(* IEC 61131-3 sources: Elmo_Master/Lasal_PRG/Elmo_EtherCAT_Test_4Axis/Class/ECAT_Master_Base (part 3) *)

#ifdef ECAT_DEBUG_EVENT_CALLBACKS
      LogError("ECAT-DEBUG: Event ECATM_EVTC_DC_DISABLED occured");
#endif

//*******************************************************************************************************************************************************
    ECATM_EVTC_ESM_DC_FAILED:
    //Error code used as argument of the ECATM_EVTC_MST_TRANS_FAILED or ECATM_EVTC_SLV_TRANS_FAILED event after the DC module failed.

#ifdef ECAT_DEBUG_EVENT_CALLBACKS
      LogError("ECAT-DEBUG: Event ECATM_EVTC_ESM_DC_FAILED occured");
#endif

//*******************************************************************************************************************************************************
    ECATM_EVTC_EOE_MBX_BAD_RSP:
    //Invalid EoE mailbox size received
    //arg1 ... slave index: int
    //arg2 ... EoE mailbox size:
    //arg3 ... EoE mailbox frame type: int

#ifdef ECAT_DEBUG_EVENT_CALLBACKS
      LogValue("ECAT-DEBUG: Invalid EoE mailbox size received. SlaveIndex: 0x{0}",evt^.arg1$UDINT);
      LogValue("ECAT-DEBUG: MBxSize: 0x{0}, MBxFrameType: 0x{1}",evt^.arg2$UDINT, evt^.arg3$UDINT);
#endif

//*******************************************************************************************************************************************************
    ECATM_EVTC_EOE_FRM_TRF_TMO:
    //Frame fragment timeout occurred. Frame was dropped
    //arg1 ... slave index: int

#ifdef ECAT_DEBUG_EVENT_CALLBACKS
      LogValue("ECAT-DEBUG: Invalid EoE mailbox size received. SlaveIndex: 0x{0}",evt^.arg1$UDINT);
#endif

//*******************************************************************************************************************************************************
    ECATM_EVTC_EOE_FRM_DROP_HDL:
    //Frame dropped because of no free frame handle available
    //arg1 ... slave index: int

#ifdef ECAT_DEBUG_EVENT_CALLBACKS
      LogValue("ECAT-DEBUG: EOE: Frame dropped because of no free frame handle available. SlaveIndex: 0x{0}",evt^.arg1$UDINT);
#endif

//*******************************************************************************************************************************************************
    ECATM_EVTC_EOE_FRM_DROP_SIZE:
    //Frame with invalid size received. Frame was dropped
    //arg1 ... slave index: int

#ifdef ECAT_DEBUG_EVENT_CALLBACKS
      LogValue("ECAT-DEBUG: EOE: Frame with invalid size received. Frame was dropped. SlaveIndex: 0x{0}",evt^.arg1$UDINT);
#endif

//*******************************************************************************************************************************************************
    ECATM_EVTC_EOE_SAT_MAC_ADD:
    //Frame with a not yet known MAC received. MAC added to switch address table
    //arg1 ... Device index: int
    //arg2 ... arg3 MAC address: arg2[3] : arg2[2] : arg2[1] : arg2[0] : arg3[1] : arg2[0]

#ifdef ECAT_DEBUG_EVENT_CALLBACKS
      LogValue("ECAT-DEBUG: EOE: Frame with a not yet known MAC received. MAC added to switch address table. DeviceIndex: 0x{0}",evt^.arg1$UDINT);
      LogValue("ECAT-DEBUG: MACADDR: 0x{0}0x{1}",evt^.arg2$UDINT, evt^.arg3$UDINT);//Before Use, should be formated correctly
#endif

//*******************************************************************************************************************************************************
    ECATM_EVTC_EOE_SAT_MAC_RM:
    //MAC is dropped from switch address table
    //arg1 ... Device index: int
    //arg2 ... arg3 MAC address: arg2[3] : arg2[2] : arg2[1] : arg2[0] : arg3[1] : arg2[0]

#ifdef ECAT_DEBUG_EVENT_CALLBACKS
      LogValue("ECAT-DEBUG: EOE: MACAddr is dropped from switch address table. DeviceIndex: 0x{0}",evt^.arg1$UDINT);
      LogValue("ECAT-DEBUG: MACADDR: 0x{0}0x{1}",evt^.arg2$UDINT, evt^.arg3$UDINT);//Before Use, should be formated correctly
#endif

//*******************************************************************************************************************************************************
    ECATM_EVTC_FRM_BAD_FRMIDX:
    // A frame with a bad index was received
    // arg1 max allowed IDX field value: int
    // arg2 received IDX field value: int

#ifdef ECAT_DEBUG_EVENT_CALLBACKS
    HWC_LogPrintf(pThis:=this, format:="@ECAT-DEBUG: A frame with a bad index was received");
    HWC_LogPrintf(pThis:=this, format:="@ECAT-DEBUG: max allowed IDX field value: %d received IDX field value: %d.", #evt^.arg1, #evt^.arg2);
#endif

//*******************************************************************************************************************************************************
    ECATM_EVTC_FRM_CFG_OP_SIZE:
    // maximal frame size during OP is too small
    // arg1 configured value (_ecatm_cfg field frmsizeop): int
    // arg2 required value: int

#ifdef ECAT_DEBUG_EVENT_CALLBACKS
    HWC_LogPrintf(pThis:=this, format:="@ECAT-DEBUG: Maximal frame size during OP is too small");
    HWC_LogPrintf(pThis:=this, format:="@ECAT-DEBUG: configured value (_ecatm_cfg field frmsizeop): %d required value: %d.", #evt^.arg1, #evt^.arg2);
#endif

//*******************************************************************************************************************************************************
    ECATM_EVTC_CRD_STATUS_CHANGED:
    // The status of the network cable redundancy diagnostics has changed
    // arg1 _ecatm_crd_status pos0 field: int
    // arg2 _ecatm_crd_status pos1 field: int
    // arg3 _ecatm_crd_status flags field: int

#ifdef ECAT_DEBUG_EVENT_CALLBACKS
    HWC_LogPrintf(pThis:=this, format:="@ECAT-DEBUG: The status of the network cable redundancy diagnostics has changed");
    HWC_LogPrintf(pThis:=this, format:="@ECAT-DEBUG: _ecatm_crd_status pos0 field: %d _ecatm_crd_status pos1 field: %d.", #evt^.arg1, #evt^.arg2);
    HWC_LogPrintf(pThis:=this, format:="@ECAT-DEBUG: _ecatm_crd_status flags field: %d", #evt^.arg3);
#endif

//*******************************************************************************************************************************************************
    ECATM_EVTC_SOE_SSC_NOTIFY:
    // SoE Notify received
    // arg1 slave index: int
    // arg2 driveno: uint8_t
    // arg3 idn: uint16_t
    // arg4 status data (16bit) from slave

#ifdef ECAT_DEBUG_EVENT_CALLBACKS
    HWC_LogPrintf(pThis:=this, format:="@ECAT-DEBUG: SoE Notify received");
    HWC_LogPrintf(pThis:=this, format:="@ECAT-DEBUG: slave index: %d driveno: uint8_t: %d.", #evt^.arg1, #evt^.arg2);
    HWC_LogPrintf(pThis:=this, format:="@ECAT-DEBUG: idn: %d status data (16bit) from slave: %d", #evt^.arg3, #evt^.arg4);
#endif

//*******************************************************************************************************************************************************
    ECATM_EVTC_SOE_SSC_TRF_TMO:
    // SoE timeout error detected
    // arg1

#ifdef ECAT_DEBUG_EVENT_CALLBACKS
    HWC_LogPrintf(pThis:=this, format:="@ECAT-DEBUG: SoE timeout error detected");
#endif

//*******************************************************************************************************************************************************
    ECATM_EVTC_SOE_SSC_TRF_ERR:
    // SoE slave responded with an error
    // arg1 slave index: int
    // arg2 driveno: uint8_t
    // arg3 idn: uint16_t
    // arg4 SoE error code from slave: uint16_t

#ifdef ECAT_DEBUG_EVENT_CALLBACKS
    HWC_LogPrintf(pThis:=this, format:="@ECAT-DEBUG: SoE slave responded with an error");
    HWC_LogPrintf(pThis:=this, format:="@ECAT-DEBUG: slave index: %d driveno: uint8_t: %d.", #evt^.arg1, #evt^.arg2);
    HWC_LogPrintf(pThis:=this, format:="@ECAT-DEBUG: idn: %d SoE error code from slave: uint16_t: %d", #evt^.arg3, #evt^.arg4);
#endif

//*******************************************************************************************************************************************************
    ECATM_EVTC_SOE_SSC_BAD_RSP:
    // Bad SoE response received
    // arg1 slave index: int

#ifdef ECAT_DEBUG_EVENT_CALLBACKS
    HWC_LogPrintf(pThis:=this, format:="@ECAT-DEBUG: Bad SoE response received. slave index: %d", #evt^.arg1);
#endif

//*******************************************************************************************************************************************************
    ECATM_EVTC_SOE_SSC_RD_BUFSIZE:
    // SoE read failed because of invalid receive buffer size
    // arg1 slave index: int
    // arg2 driveno: uint8_t
    // arg3 idn: uint16_t
    // arg4 required size: int

#ifdef ECAT_DEBUG_EVENT_CALLBACKS
    HWC_LogPrintf(pThis:=this, format:="@ECAT-DEBUG: SoE read failed because of invalid receive buffer size");
    HWC_LogPrintf(pThis:=this, format:="@ECAT-DEBUG: slave index: %d driveno: uint8_t: %d.", #evt^.arg1, #evt^.arg2);
    HWC_LogPrintf(pThis:=this, format:="@ECAT-DEBUG: idn: %d required size: %d", #evt^.arg3, #evt^.arg4);
#endif

//*******************************************************************************************************************************************************
    ECATM_EVTC_SOE_SSC_RD_FRAG:
    // SoE read failed because of unexpected fragment number
    // arg1 slave index: int
    // arg2 driveno: uint8_t
    // arg3 idn: uint16_t

#ifdef ECAT_DEBUG_EVENT_CALLBACKS
    HWC_LogPrintf(pThis:=this, format:="@ECAT-DEBUG: SoE read failed because of unexpected fragment number");
    HWC_LogPrintf(pThis:=this, format:="@ECAT-DEBUG: slave index: %d driveno: uint8_t: %d.", #evt^.arg1, #evt^.arg2);
    HWC_LogPrintf(pThis:=this, format:="@ECAT-DEBUG: idn: %d.", #evt^.arg3);
#endif

//*******************************************************************************************************************************************************
    ECATM_EVTC_SII_EEPROM_BUSY_TMO:
    // SII EEPROM access failed because of EEPROM busy flag
    // arg1 slave index: int
    // arg2 SII Status Register (ESC register 0x502): uint8_t

#ifdef ECAT_DEBUG_EVENT_CALLBACKS
    HWC_LogPrintf(pThis:=this, format:="@ECAT-DEBUG: SII EEPROM access failed because of EEPROM busy flag");
    HWC_LogPrintf(pThis:=this, format:="@ECAT-DEBUG: slave index: %d SII Status Register (ESC register 0x502): uint8_t: %x.", #evt^.arg1, #evt^.arg2);
#endif

//*******************************************************************************************************************************************************
    ECATM_EVTC_SII_EEPROM_PDI_TMO:
    // SII EEPROM access failed as owenership is with PDI
    // arg1 slave index: int

#ifdef ECAT_DEBUG_EVENT_CALLBACKS
    HWC_LogPrintf(pThis:=this, format:="@ECAT-DEBUG: SII EEPROM access failed as owenership is with PDI. slave index: %d", #evt^.arg1);
#endif

//*******************************************************************************************************************************************************
    ECATM_EVTC_SII_INVALID_VERSION:
    // SII read till end failed as SII version is invalid
    // arg1 slave index: int
    // arg2 SII version field (0x3F) (should be 0x001): uint16_t

#ifdef ECAT_DEBUG_EVENT_CALLBACKS
    HWC_LogPrintf(pThis:=this, format:="@ECAT-DEBUG: SII read till end failed as SII version is invalid");
    HWC_LogPrintf(pThis:=this, format:="@ECAT-DEBUG: slave index: %d SII version field (0x3F) (should be 0x001): %x.", #evt^.arg1, #evt^.arg2);
#endif

//*******************************************************************************************************************************************************
    ECATM_EVTC_HC_TOO_MANY_DEVICES:
    // The number of found devices during HC detection exceeds the number of devices defined in the ENI
    // arg1 found devices: int
    // arg2 number of devices in ENI: int

#ifdef ECAT_DEBUG_EVENT_CALLBACKS
    HWC_LogPrintf(pThis:=this, format:="@ECAT-DEBUG: The number of found devices during HC detection exceeds the number of devices defined in the ENI");
    HWC_LogPrintf(pThis:=this, format:="@ECAT-DEBUG: found devices: %d number of devices in ENI: %d.", #evt^.arg1, #evt^.arg2);
#endif

//*******************************************************************************************************************************************************
    ECATM_EVTC_HC_GRP_SEARCH:
    // Start searching for matching HC group connected to a device port
    // arg1 slave index: int
    // arg2 port index: enum {ECAT_ESC_PORT_A; ECAT_ESC_PORT_B; ECAT_ESC_PORT_C; ECAT_ESC_PORT_D}

#ifdef ECAT_DEBUG_EVENT_CALLBACKS
    HWC_LogPrintf(pThis:=this, format:="@ECAT-DEBUG: Start searching for matching HC group connected to a device port");
    HWC_LogPrintf(pThis:=this, format:="@ECAT-DEBUG: slave index: %d port index: %d.", #evt^.arg1, #evt^.arg2);
#endif

//*******************************************************************************************************************************************************
    ECATM_EVTC_HC_GRP_FOUND:
    // Found a matching HC group connected to the device port
    // arg1 HC group index matching: int
    // arg2 slave index: int
    // arg3 port index: enum {ECAT_ESC_PORT_A; ECAT_ESC_PORT_B; ECAT_ESC_PORT_C; ECAT_ESC_PORT_D}

#ifdef ECAT_DEBUG_EVENT_CALLBACKS
    HWC_LogPrintf(pThis:=this, format:="@ECAT-DEBUG: Found a matching HC group connected to the device port");
    HWC_LogPrintf(pThis:=this, format:="@ECAT-DEBUG: HC group index that is no longer reachable: %d.", #evt^.arg1);
    HWC_LogPrintf(pThis:=this, format:="@ECAT-DEBUG: slave index: %d port index: %d.", #evt^.arg2, #evt^.arg3);
#endif

//*******************************************************************************************************************************************************
    ECATM_EVTC_HC_GRP_NO_MATCH:
    // Failed to find a matching HC group for the device port
    // arg1 slave index: int
    // arg2 port index: enum {ECAT_ESC_PORT_A; ECAT_ESC_PORT_B; ECAT_ESC_PORT_C; ECAT_ESC_PORT_D}

#ifdef ECAT_DEBUG_EVENT_CALLBACKS
    HWC_LogPrintf(pThis:=this, format:="@ECAT-DEBUG: Failed to find a matching HC group for the device port");
    HWC_LogPrintf(pThis:=this, format:="@ECAT-DEBUG: slave index: %d port index: %d.", #evt^.arg1, #evt^.arg2);
#endif

//*******************************************************************************************************************************************************
    ECATM_EVTC_HC_GRP_DISCONNECTED:
    // Hot Connect group is disconnected from the device port
    // arg1 HC group index that is no longer reachable: int
    // arg2 slave index: int
    // arg3 port index: enum {ECAT_ESC_PORT_A; ECAT_ESC_PORT_B; ECAT_ESC_PORT_C; ECAT_ESC_PORT_D}

#ifdef ECAT_DEBUG_EVENT_CALLBACKS
    HWC_LogPrintf(pThis:=this, format:="@ECAT-DEBUG: Hot Connect group is disconnected from the device port");
    HWC_LogPrintf(pThis:=this, format:="@ECAT-DEBUG: HC group index that is no longer reachable: %d.", #evt^.arg1);
    HWC_LogPrintf(pThis:=this, format:="@ECAT-DEBUG: slave index: %d port index: %d.", #evt^.arg2, #evt^.arg3);
#endif

//*******************************************************************************************************************************************************
    ECATM_EVTC_HC_PORT_CHANGED:
    // The status of device port has changed
    // arg1 slave index: int
    // arg2 port index: enum {ECAT_ESC_PORT_A; ECAT_ESC_PORT_B; ECAT_ESC_PORT_C; ECAT_ESC_PORT_D}
    // arg3 new status: flags see ECATM_HC_PORT_FLAG…
    // arg4 old status: flags see ECATM_HC_PORT_FLAG…

#ifdef ECAT_DEBUG_EVENT_CALLBACKS
    HWC_LogPrintf(pThis:=this, format:="@ECAT-DEBUG: The status of device port has changed");
    HWC_LogPrintf(pThis:=this, format:="@ECAT-DEBUG: slave index: %d port index: %d.", #evt^.arg1, #evt^.arg2);
    HWC_LogPrintf(pThis:=this, format:="@ECAT-DEBUG: new status: %d old status: %d.", #evt^.arg3, #evt^.arg4);
#endif

//*******************************************************************************************************************************************************
    ECATM_EVTC_HC_PORT_OPEN:
    // A device port will be opened to connect new devices
    // arg1 slave index: int
    // arg2 port index: enum {ECAT_ESC_PORT_A; ECAT_ESC_PORT_B; ECAT_ESC_PORT_C; ECAT_ESC_PORT_D}

#ifdef ECAT_DEBUG_EVENT_CALLBACKS
    HWC_LogPrintf(pThis:=this, format:="@ECAT-DEBUG: A device port will be opened to connect new devices");
    HWC_LogPrintf(pThis:=this, format:="@ECAT-DEBUG: slave index: %d port index: %d.", #evt^.arg1, #evt^.arg2);
#endif

//*******************************************************************************************************************************************************
    ECATM_EVTC_HC_MAN_PORT_CLOSED:
    // A mandatory connection at the device port is closed/disconnected
    // arg1 slave index: int
    // arg2 port index: enum {ECAT_ESC_PORT_A; ECAT_ESC_PORT_B; ECAT_ESC_PORT_C; ECAT_ESC_PORT_D}

#ifdef ECAT_DEBUG_EVENT_CALLBACKS
    HWC_LogPrintf(pThis:=this, format:="@ECAT-DEBUG: A mandatory connection at the device port is closed/disconnected");
    HWC_LogPrintf(pThis:=this, format:="@ECAT-DEBUG: slave index: %d port index: %d.", #evt^.arg1, #evt^.arg2);
#endif

//*******************************************************************************************************************************************************
    ECATM_EVTC_HC_MAN_PORT_OPENING:
    // Opening a connection at the device port which is closed
    // arg1 slave index: int
    // arg2 port index: enum {ECAT_ESC_PORT_A; ECAT_ESC_PORT_B; ECAT_ESC_PORT_C; ECAT_ESC_PORT_D}

#ifdef ECAT_DEBUG_EVENT_CALLBACKS
    HWC_LogPrintf(pThis:=this, format:="@ECAT-DEBUG: Opening a connection at the device port which is closed");
    HWC_LogPrintf(pThis:=this, format:="@ECAT-DEBUG: slave index: %d port index: %d.", #evt^.arg1, #evt^.arg2);
#endif

//*******************************************************************************************************************************************************
    ECATM_EVTC_HC_TOPO_INVALID:
    // The Hot Connect topology solver failed to match the current network topology

#ifdef ECAT_DEBUG_EVENT_CALLBACKS
    HWC_LogPrintf(pThis:=this, format:="@ECAT-DEBUG: The Hot Connect topology solver failed to match the current network topology");
#endif

//*******************************************************************************************************************************************************
    ECATM_EVTC_HC_SLV_NOT_CONNECTED:
    // The current device is part of a not connected HC group

#ifdef ECAT_DEBUG_EVENT_CALLBACKS
    HWC_LogPrintf(pThis:=this, format:="@ECAT-DEBUG: The current device is part of a not connected HC group");
#endif

//*******************************************************************************************************************************************************
    ECATM_EVTC_DC_PROPDLY_UPDATE:
    // The Distributed Clocks module is starting an propagation delay update run
    // The force flag is set when not triggered via _ecatm_dc_cfg.propdly_update_ms timeout.
    // arg1 forced run: bool

#ifdef ECAT_DEBUG_EVENT_CALLBACKS
    HWC_LogPrintf(pThis:=this, format:="@ECAT-DEBUG: The Distributed Clocks module is starting an propagation delay update run");
    HWC_LogPrintf(pThis:=this, format:="@ECAT-DEBUG: The force flag is set when not triggered via _ecatm_dc_cfg.propdly_update_ms timeout. forced run: %d", #evt^.arg1);
#endif

//*******************************************************************************************************************************************************
    ECATM_EVTC_DC_PROPDLY_FINISHED:
    // The propagation delay is now updated

#ifdef ECAT_DEBUG_EVENT_CALLBACKS
    HWC_LogPrintf(pThis:=this, format:="@ECAT-DEBUG: The propagation delay is now updated");
#endif

//*******************************************************************************************************************************************************
    ECATM_EVTC_DC_SLV_SYNC_TIMOUT:
    // The static drift compensation for a single device during during operation failed
    // arg1 slave index: int
    // arg2 last syncwin measured: unsigned int

#ifdef ECAT_DEBUG_EVENT_CALLBACKS
    HWC_LogPrintf(pThis:=this, format:="@ECAT-DEBUG: The static drift compensation for a single device during during operation failed");
    HWC_LogPrintf(pThis:=this, format:="@ECAT-DEBUG: slave index: %d last syncwin measured: %d.", #evt^.arg1, #evt^.arg2);
#endif

//*******************************************************************************************************************************************************
    ECATM_EVTC_FOE_ERROR_RSP:
    // Error code set by FoE, when an error response was received or send via ECATM_FOE_REQ_ERROR.
#ifdef ECAT_DEBUG_EVENT_CALLBACKS
    HWC_LogPrintf(pThis:=this, format:="@ECAT-DEBUG: Error code set by FoE, when an error response was received or send via ECATM_FOE_REQ_ERROR");
#endif

//*******************************************************************************************************************************************************
    ECATM_EVTC_FOE_USER_ABORT:
    // Error code set by FoE, when FoE transfer was aborted by a user request.
#ifdef ECAT_DEBUG_EVENT_CALLBACKS
    HWC_LogPrintf(pThis:=this, format:="@ECAT-DEBUG: Error code set by FoE, when FoE transfer was aborted by a user request");
#endif

//*******************************************************************************************************************************************************
    ECATM_EVTC_FOE_UNEXP_RSP:
    // Warning generated when an unexpected unhandled FoE mbx message is received.
    // This could be a followup of an abort or error.
    // arg1 slave index: int
    // arg2 opcode Byte[0] of msg: uint8_t
    // arg3 length of FoE the message excluding the mbx header: int
#ifdef ECAT_DEBUG_EVENT_CALLBACKS
    HWC_LogPrintf(pThis:=this, format:="@ECAT-DEBUG: Warning generated when an unexpected unhandled FoE mbx message is received");
    HWC_LogPrintf(pThis:=this, format:="@ECAT-DEBUG: slave index: %d opcode Byte[0] of msg: %V1.", #evt^.arg1, #evt^.arg2);
    HWC_LogPrintf(pThis:=this, format:="@ECAT-DEBUG: length of FoE the message excluding the mbx header: %d.", #evt^.arg3);
#endif

//*******************************************************************************************************************************************************
    ECATM_EVTC_MBX_WR_PROT_FAILED:
    // Mailbox write request failed. New event combining all mailbox protocol related write errors.
    // arg1 slave index: int
    // arg2 The mailbox protocol (ECAT_MBX_TYPE…): uint8_t
    // arg3 The mailbox error reason (lower layer): int
#ifdef ECAT_DEBUG_EVENT_CALLBACKS
    HWC_LogPrintf(pThis:=this, format:="@ECAT-DEBUG: Mailbox write request failed. New event combining all mailbox protocol related write errors");
    HWC_LogPrintf(pThis:=this, format:="@ECAT-DEBUG: slave index: %d The mailbox protocol (ECAT_MBX_TYPE…): %V1.", #evt^.arg1, #evt^.arg2);
    HWC_LogPrintf(pThis:=this, format:="@ECAT-DEBUG: The mailbox error reason (lower layer): %d.", #evt^.arg3);
#endif

//*******************************************************************************************************************************************************
    ECATM_EVTC_ESM_INVALID_WKC_SO:
    // The working counter check during SafeOP hit a timeout. This can happen for some devices that do not handle outputs or inputs correctly during SafeOP.
    // The ecat master continues in this case after a timeout with this warning.
    // arg1 cyclic task idx: int (index of cyclic task with invalid WKC)
#ifdef ECAT_DEBUG_EVENT_CALLBACKS
    HWC_LogPrintf(pThis:=this, format:="@ECAT-DEBUG: The WKC check during SafeOP hit a timeout. This can happen for some devices that do not handle outputs or inputs correctly during SafeOP.");
    HWC_LogPrintf(pThis:=this, format:="@ECAT-DEBUG: cyclic task idx: int (index of cyclic task with invalid WKC): %d.", #evt^.arg1);
#endif

//*******************************************************************************************************************************************************
    ECATM_EVTC_SDOINFO_BAD_RESPONE:
    // A SDO info response with a bad length was received
    // arg1 slave index: int
    // arg2 Length of the bad response: int
#ifdef ECAT_DEBUG_EVENT_CALLBACKS
    HWC_LogPrintf(pThis:=this, format:="@ECAT-DEBUG: MA SDO info response with a bad length was received");
    HWC_LogPrintf(pThis:=this, format:="@ECAT-DEBUG: slave index: %d Length of the bad response:: %d.", #evt^.arg1, #evt^.arg2);
#endif

//*******************************************************************************************************************************************************
    ECATM_EVTC_SDOINFO_UNEXP:
    // A valid SDO info response/request was received but no waiting handle is attached
    // arg1 slave index: int
    // arg2 SdoInfo opcode: uint8_t
    // arg3 Length of the bad response: int
#ifdef ECAT_DEBUG_EVENT_CALLBACKS
    HWC_LogPrintf(pThis:=this, format:="@ECAT-DEBUG: A valid SDO info response/request was received but no waiting handle is attached");
    HWC_LogPrintf(pThis:=this, format:="@ECAT-DEBUG: slave index: %d SdoInfo opcode: %V1.", #evt^.arg1, #evt^.arg2);
    HWC_LogPrintf(pThis:=this, format:="@ECAT-DEBUG: Length of the bad response: %d.", #evt^.arg3);
#endif

//*******************************************************************************************************************************************************
    ECATM_EVTC_SDOINFO_BAD_FRG:
    // Received a unexpected and bad fragment number
    // arg1 slave index: int
    // arg2 fragleft received: int
    // arg3 fragleft expected: int
#ifdef ECAT_DEBUG_EVENT_CALLBACKS
    HWC_LogPrintf(pThis:=this, format:="@ECAT-DEBUG: Received a unexpected and bad fragment number");
    HWC_LogPrintf(pThis:=this, format:="@ECAT-DEBUG: slave index: %d", #evt^.arg1);
    HWC_LogPrintf(pThis:=this, format:="@ECAT-DEBUG: ragleft received: %d. fragleft expected: %d", #evt^.arg2, #evt^.arg3);
#endif

//*******************************************************************************************************************************************************
    ECATM_EVTC_SDOINFO_EMPTY:
    // Return code only. The error is set when an SDO info transfer is succeeded without any payload was received.
    // This is a workaround for the SSC which can be seen when a transfer is aborted through a INIT transition.
#ifdef ECAT_DEBUG_EVENT_CALLBACKS
    HWC_LogPrintf(pThis:=this, format:="@ECAT-DEBUG: The error is set when an SDO info transfer is succeeded without any payload was received.");
#endif

  end_case;

END_FUNCTION

FUNCTION __CDECL VIRTUAL ECAT_Master_Base::SendEvtCallBacktoSlave
	VAR_INPUT
		udMasterID 	: UDINT;
		evt 	: ^t_st_ecatm_evt;
		EventType 	: DINT;
		uiCallbackInfo 	: UINT;
	END_VAR
  VAR
    pCurrentSlave : ^t_sSlaveInfo;
    _Para 	  : CmdStruct;
    _Result 	: Results;
    ret_code 	: IprStates;
  END_VAR

  // INFO_CALLBACK: Callbacks may be received immediately after setting the callback method because EtherCAT Master may run on a different core!
  // INFO_CALLBACK: As of 15.07. Slave callback (search for SendEvtCallBacktoSlave) are not called until the first call to OS_ECATM_MST_REQ_STATE in the PostInit.
  // INFO_CALLBACK: This guarantees that the data structure needed in SendEvtCallBacktoSlave are initialized, before the 1st callback is received.

  //Check if we got a valid slave number
  if evt^.arg1$UDINT <= sSlaveInfo.udMaxSlaves then

    pCurrentSlave := sSlaveInfo.pSlaves + (evt^.arg1$UDINT * sizeof(t_sSlaveInfo)); //Set pointer to correct slave

    if (pCurrentSlave) & (pCurrentSlave^.pThis) then

      _Para.uiCmd                     := ECAT_M_EVENT_CALLBACK;
      _Para.aPara[0]                  := 1;
      _Para.aPara[1]$UDINT            := udMasterID;
      _Para.aPara[2]$^t_st_ecatm_evt  := evt;
      _Para.aPara[3]                  := EventType;
      _Para.aPara[4]                  := uiCallbackInfo;

      //Forward event callback via newinst to respective Slave
      ret_code := pCurrentSlave^.pThis^.NewInst(#_Para,#_Result);

      if (ret_code <> READY) |(_Result.uiLng <> 8) |
         (_Result.aData[0]$DINT <> ECAT_RETOK) |
         (_Result.aData[4]$DINT <> 1) then // Version

        if (uiCallbackInfo = LSL_ECATM_ACYCLIC_TASK) then
          LogValue("@0577 (ECAT_Master_Base::SendEvtCallBacktoSlave) NewInstCmd: ECAT_M_EVENT_CALLBACK Failed! ret_code = 0x{0}, return code = 0x{1}, Version = 0x{2}", ret_code$UDINT, _Result.aData[0]$UDINT, _Result.aData[4]$UDINT);
        else
          bd_LogRtMessagesInCy.PostIt.SendEvtCallInvFailed := TRUE;
          bd_LogRtMessagesInCy.aLogValue1[7] := _Result.aData[0]$UDINT;
        end_if;

      end_if;
    end_if;
  else

    if (uiCallbackInfo = LSL_ECATM_ACYCLIC_TASK) then
      LogValue("@0576 (ECAT_Master_Base::SendEvtCallBacktoSlave) Invalid slave number from Event callback! evt^.arg1 = 0x{0}, sSlaveInfo.udMaxSlaves = 0x{1}, Event: 0x{2}", evt^.arg1$UDINT, sSlaveInfo.udMaxSlaves, evt^.evtcode$UDINT);
    else
      bd_LogRtMessagesInCy.PostIt.SendEvtCallInvSlv := TRUE;
      bd_LogRtMessagesInCy.aLogValue1[6] := evt^.arg1$UDINT;
    end_if;

  end_if;

END_FUNCTION

FUNCTION VIRTUAL ECAT_Master_Base::SetRequiredError
	VAR_INPUT
		pTargetThis 	: ^ECAT_Slave_Base;(* := NIL *)
		udSlaveIndex 	: UDINT;(* := 16#FFFFFFFF *)
		bLogInMethAllowed 	: BOOL;(* := FALSE *)
	END_VAR

  if pTargetThis & udSlaveIndex <> 16#FFFFFFFF then
    pTargetThis^.ClassState := _RequiredError;

    if bLogInMethAllowed then
      LogValue("@0579 (ECAT_Master_Base::SetRequiredError) Required Error on EtherCAT Slave 0x{0}.", udSlaveIndex);
    else
      bd_LogRtMessagesInCy.PostIt.SetReqErrSlv := TRUE;
      bd_LogRtMessagesInCy.aLogValue1[8] := udSlaveIndex;
    end_if;

  else

    // general required error (initialisation failed)
    // if no required module => don't crash
    if (bd_Flags.bIsRequired = FALSE) then
      return;
    end_if;

  end_if;

  ClassState := _RequiredError;

  //Set off the HardwareControl class
  ToHwControl.SetHardwareOff(e_error:=_RequiredError);

  if pECAT then
    // if a required module is not available or doesn't work properly, the system should crash
    OS_ECATM_raise_error(pECAT,0,"Required Error");
  else

    if bLogInMethAllowed then
      LogError("@057A (ECAT_Master_Base::SetRequiredError) Failed to raise Required Error.");
    else
      bd_LogRtMessagesInCy.PostIt.SetReqErrFailed := TRUE;
    end_if;

  end_if;

END_FUNCTION

#pragma warning(disable:73);
FUNCTION VIRTUAL ECAT_Master_Base::ConnectEvent
	VAR_INPUT
		udMasterID 	: UDINT;
		evt 	: ^t_st_ecatm_evt;
		EventType 	: DINT;
		uiCallbackInfo 	: UINT;
	END_VAR

  InitSSW := _StartInit;

  //      OS_ECATM_MST_REQ_STATE(pECAT, ecatmhdl, (ECAT_STATE_OP)$UDINT , StateTransitionBehaviour);

END_FUNCTION
#pragma warning(default:73);

FUNCTION VIRTUAL ECAT_Master_Base::DisconnectEvent
	VAR_INPUT
		udMasterID 	: UDINT;
		evt 	: ^t_st_ecatm_evt;
		EventType 	: DINT;
		uiCallbackInfo 	: UINT;
	END_VAR
  VAR
  	pCurrentSlave : ^t_sSlaveInfo;
    i : UDINT;
  END_VAR

  if (InitSSW <> _InitFinished) &
     (InitSSW <> _PrepareError) &
     (InitSSW <> _ErrorOccured)  then
    return;
  end_if;

  InitSSW := _NotConnected;
  udDisconnectEventTime := ops.tAbsolute;

  // if there is a required error, we would disguise it, if we call the disconnect interfaces
  if ClassState <> _RequiredError then

    // tell all the connected modules
    if sSlaveInfo.udMaxSlaves then
      pCurrentSlave := sSlaveInfo.pSlaves; //Point to current slave
      for i:=0 to sSlaveInfo.udMaxSlaves-1 do
        if pCurrentSlave^.pThis then
          pCurrentSlave^.pThis^.DisconnectEvent();
        end_if;
        pCurrentSlave += sizeof(t_sSlaveInfo);
      end_for;
    end_if;
  end_if;

END_FUNCTION

FUNCTION VIRTUAL GLOBAL ECAT_Master_Base::GetFrameTimesPointer
	VAR_INPUT
		udCycTaskID 	: UDINT;
	END_VAR
	VAR_OUTPUT
		pEtherCATFrameTimes 	: ^t_s_EtherCATFrameTimes;
	END_VAR

  pEtherCATFrameTimes := NIL;

  //Check for valid Task ID
  if udNoCycTasks & pCycTaskInfo then
    if udCycTaskID > udNoCycTasks-1 then
      return; // Return default NIL
    end_if;

    pEtherCATFrameTimes := #pCycTaskInfo^.sFrameTimes + ( sizeof(t_s_CycTaskInfo) * udCycTaskID);
  end_if;

END_FUNCTION

FUNCTION VIRTUAL ECAT_Master_Base::GetPointer2ObjectPath
	VAR_OUTPUT
		p_us_ObjectPath 	: ^USINT;
	END_VAR

  if pObjectPath = NIL then
    // create object path for the PLC
    aObjectPath[0] := 2;    // pObjectPath uses 1 Byte length and one Byte Domain
    aObjectPath[1] := 0;
    aObjectPath[2] := HWT_ESCAPE_ECAT;

    pObjectPath := #aObjectPath[0];
  end_if;

  p_us_ObjectPath := pObjectPath;

END_FUNCTION

FUNCTION VIRTUAL ECAT_Master_Base::GetCallInitModuleTimeout
	VAR_OUTPUT
		udTimeout 	: UDINT;
	END_VAR

  //Method can be overwritten if standard timeout is too high/too less for application
  udTimeout := ECATM_INIT_CALLINITMODULE_TIMEOUT;

END_FUNCTION

FUNCTION VIRTUAL ECAT_Master_Base::GetWait4SynchronTimeout
	VAR_OUTPUT
		udTimeout 	: UDINT;
	END_VAR

  //Method can be overwritten if standard timeout is too high/too less for application
  udTimeout := ECATM_WAIT_FOR_SYNCHRON_TIMEOUT;

END_FUNCTION

FUNCTION VIRTUAL ECAT_Master_Base::GetWait4LinkTimeout
	VAR_OUTPUT
		udTimeout 	: UDINT;
	END_VAR

  //Method can be overwritten if standard timeout is too high/too less for application
  udTimeout := ECATM_INIT_LINK_TIMEOUT;

END_FUNCTION

FUNCTION VIRTUAL ECAT_Master_Base::ProcessFrameErrorCheck
	VAR_INPUT
		udPrcstate 	: UDINT;
	END_VAR
	VAR_OUTPUT
		dTriggerFrameError 	: DINT;
	END_VAR

  dTriggerFrameError := 1;

  aFrameErrorLogBuffer[udCurrentLogEntry].udTimeStamp     := ops.tAbsolute;
  aFrameErrorLogBuffer[udCurrentLogEntry].bdProcessState  := udPrcstate$BDINT;

  udCurrentLogEntry += 1;

  //Check for array limit
  if udCurrentLogEntry > ECATM_MAX_SIZE_FRAME_ERROR_LOGBUFFER-1 then
    udCurrentLogEntry := 0;
  end_if;

  //It is possible and allowed that sometimes a frame is missing. With this check the user can set how many consecutive missing frames
  //are going to raise an error.
  sDebugCounters.udConsecutiveMissingFrameCounter += 1;
  sDebugCounters.udTotalMissingFrameCounter += 1;

  case MissingFrameBehaviour of

    0 : dTriggerFrameError := 0;  //If dTriggerFrameError is zero, no error will be raised and the application will work with the data from the last valid frame/cycle
                                  //Do not trigger an error due to client setting

    1 : dTriggerFrameError := 1;   //trigger an error due to client setting

    else
      //Check for number of missing frames and client setting
      if MissingFrameBehaviour > sDebugCounters.udConsecutiveMissingFrameCounter  then
        dTriggerFrameError := 0;  //no error due to client setting
      end_if;
  end_case;

END_FUNCTION

FUNCTION VIRTUAL ECAT_Master_Base::ExtendPostInitTime
	VAR_INPUT
		AdditionalTime 	: UDINT;
	END_VAR
  VAR
  	MyPara          : CmdStruct;
    MyResult        : results;
  END_VAR

  MyPara.uiCmd    := CMD_EXTEND_POST_INIT_TIME;
  MyPara.aPara[0] := AdditionalTime$DINT;

  if ToHwControl.NewInst(#MyPara, #MyResult) <> READY then
    // Just log, default Postinit may be enough anyway. Otherwise it will timeout in postinit.
    LogValue("@084B (ECAT_Master_Base::ExtendPostInitTime) Failed to increase Postinit-Timeout by 0x{0}.", AdditionalTime);
  end_if;

END_FUNCTION

FUNCTION VIRTUAL ECAT_Master_Base::SendManagerErrorToSlaves
  VAR
    pCurrentSlave : ^t_sSlaveInfo;
    i             : UDINT;
  	MyPara          : CmdStruct;
    MyResult        : results;
  END_VAR

  pCurrentSlave := sSlaveInfo.pSlaves; //Point to current slave

  MyPara.uiCmd     := ECAT_M_SET_CLASSSTATE;
  MyPara.aPara[0]  := 1; // Version

  //Call Update all logged in slaves
  for i:=0 to sSlaveInfo.udMaxSlaves-1 do

    //Check if slave can be called
    if pCurrentSlave^.pThis then
      if pCurrentSlave^.pThis^.ClassState = _ClassOk then
        MyPara.aPara[1]$t_e_VaranErrors := _ManagerError;  // ClassState
      else
        // Do not overwrite already existing error state on client
        MyPara.aPara[1]$t_e_VaranErrors := pCurrentSlave^.pThis^.ClassState; // ClassState
      end_if;

      MyPara.aPara[2]$DINT := 0; // Online

      pCurrentSlave^.pThis^.NewInst(#MyPara, #MyResult);

    end_if;

    pCurrentSlave += sizeof(t_sSlaveInfo);
  end_for;

END_FUNCTION

FUNCTION VIRTUAL GLOBAL ECAT_Master_Base::DisableInitBusTimeouts
	VAR_INPUT
		AllTimeouts 	: BOOL;(* := TRUE *)
		Wait4LinkTimeOut 	: BOOL;(* := FALSE *)
		StateTransitionTimeout 	: BOOL;(* := FALSE *)
		InitModuleTimeOut 	: BOOL;(* := FALSE *)
		WaitForSynchronTimeOut 	: BOOL;(* := FALSE *)
		PostInitTimeout 	: BOOL;(* := FALSE *)
	END_VAR

  if Alltimeouts then

    bd_Flags.bDisableWait4LinkTimeOut       := TRUE;
    bd_Flags.bDisableStateTransitionTimeout := TRUE;
    bd_Flags.bDisableInitModuleTimeOut      := TRUE;
    bd_Flags.bDisableWaitForSynchronTimeOut := TRUE;
    bd_Flags.bPostInitCancel                := TRUE;

  else

    bd_Flags.bDisableWait4LinkTimeOut       := Wait4LinkTimeOut;
    bd_Flags.bDisableStateTransitionTimeout := StateTransitionTimeout;
    bd_Flags.bDisableInitModuleTimeOut      := InitModuleTimeOut;
    bd_Flags.bDisableWaitForSynchronTimeOut := WaitForSynchronTimeOut;
    bd_Flags.bPostInitCancel                := PostInitTimeout;

  end_if;

END_FUNCTION

FUNCTION VIRTUAL GLOBAL ECAT_Master_Base::DisableRequiredError
	VAR_OUTPUT
		retval 	: DINT;
	END_VAR

  retval := -1;

  if us_InitCnt <= 1 then
    bd_Flags.bDisableRequired := TRUE;
    retval := 0;
  end_if;

END_FUNCTION
